// TIA Portal V21 export
// export: Created 2026-08-21T20:18:51.5514905Z, ExportSetting None, DisplayName Totally Integrated Automation Portal, DisplayVersion V21, DisplayName STEP 7 Professional, DisplayVersion V21, DisplayName STEP 7 Safety, DisplayVersion V21, DisplayName Tech WebApplication, DisplayVersion V21, DisplayName WinCC Basic/Comfort/Advanced, DisplayVersion V21, DisplayName WinCC Professional, DisplayVersion V21, DisplayName WinCC Unified, DisplayVersion V21
DATA_BLOCK "CalcDoseDB"   // DB6
// stored: InstanceOfName CalcDose, InstanceOfType FB
"CalcDose"
   // VAR_INPUT
   //    Enable : Bool;
   //    Dose_Liters : Real;
   //    VolumeFlow : Real;
   //    Adj_high : Real;
   //    Adj_middle : Real;
   //    Adj_low : Real;
   //    Adj_high_Value : Real;
   //    Adj_middle_Value : Real;
   //    Adj_low_Value : Real;
   //    Scale_Raw : "ScaVal_Raw";
   // END_VAR
   // VAR_OUTPUT
   //    Service_Done : Bool;
   //    PIDCtrl_Value : "AnaVal";
   //    Liters { ExternalWritable := 'False'} : Real;
   //    Liters_Raw : Int;
   // END_VAR
BEGIN
END_DATA_BLOCK
